// Mitsubishi GX Works2 project: Task2_Ex_5   PLC: FX3G

PROGRAM MAIN
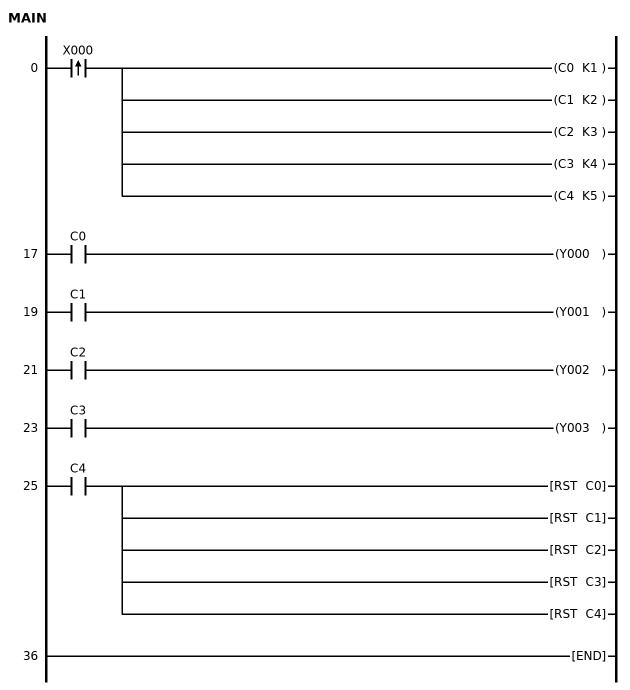
0     LDP     X000
      OUT     C0 K1
      OUT     C1 K2
      OUT     C2 K3
      OUT     C3 K4
      OUT     C4 K5
17    LD      C0
      OUT     Y000
19    LD      C1
      OUT     Y001
21    LD      C2
      OUT     Y002
23    LD      C3
      OUT     Y003
25    LD      C4
      RST     C0
      RST     C1
      RST     C2
      RST     C3
      RST     C4
36    END
END_PROGRAM
